// TIA Portal project "MoreLanguages" (V21)

(* hardware
DEVICE "PLC_Classic"  S7-300 station
   slot 0: "Rail_0"  Rail  6ES7 390-1***0-0AA0
   slot 2: "PLC_Classic"  CPU 315-2 PN/DP  6ES7 315-2EH14-0AB0  V3.2.18
      slot 2: "PROFINET interface_1"  PN-IO
         slot 1: "Port_1"  Port
         slot 2: "Port_2"  Port
DEVICE "PLC_More"  S7-1500 station
   slot 0: "Rail_0"  Rack  6ES7 590-1***0-0AA0
   slot 1: "PLC_More"  CPU 1516-3 PN/DP  6ES7 516-3AN02-0AB0  V2.9
      slot 3: "CPU display_1"  6ES7591-1BA00-0AA0
      slot 32768: "PROFINET interface_1"  X1
         slot 32769: "Port_1"  X1 P1
         slot 32770: "Port_2"  X1 P2
      slot 33024: "PROFINET interface_2"  X2
         slot 33025: "Port_1"  X2 P1
      slot 33280: "DP interface_1"  X3
      slot 34817: "Virtual CP interface port_1"  Virtual CP interface port  Virtual CP interface port
*)

// ===== PLC "PLC_Classic"  CPU 315-2 PN/DP =====

VAR_GLOBAL   // PLC tag table "Default tag table"
   "Tag__639308646888752274" AT %T1 : Timer;
   "Tag__639308646889222918" AT %I0.2 : Bool;
   "Tag__639308646889222919" AT %C1 : Counter;
   "Tag__639308646889222920" AT %I0.3 : Bool;
   "Tag__639308646889546626" AT %MW10 : Word;
   "Tag__639308646889705153" AT %QW0 : Word;
END_VAR

VAR_GLOBAL   // PLC tag table "IO"
   "Start" AT %I0.0 : Bool;   // Start button
   "Stop" AT %I0.1 : Bool;   // Stop button
   "Motor" AT %Q0.0 : Bool;   // Motor contactor
   "Raw" AT %IW2 : Int;   // Raw level
END_VAR

TYPE "Recipe"
   STRUCT
      amount : Int := 10;   // Units per batch
      heat : Bool;   // Whether the batch is heated
      dwell : Time := T#5S;   // Time in the heater
   END_STRUCT;
END_TYPE

DATA_BLOCK "Store"   // DB1
TITLE = Shared data
{ S7_Optimized_Access := 'FALSE' }
VERSION : 0.1
// A shared data block of a classic CPU, which has standard access only.
   VAR
      count : Int := 3;   // Batches made
      level : Word;
      current : "Recipe";
      flags : Array[0..7] of Bool;
   END_VAR
BEGIN
   current.amount := 12;
END_DATA_BLOCK

DATA_BLOCK "ScaleDb"   // DB2
{ S7_Optimized_Access := 'FALSE' }
VERSION : 0.1
// stored: InstanceOfName Scale
"Scale"
BEGIN
END_DATA_BLOCK

FUNCTION_BLOCK "Scale"   // FB1, SCL
TITLE = Scale a raw value
{ S7_Optimized_Access := 'FALSE' }
VERSION : 0.1
// SCL on a classic CPU.
   VAR_INPUT
      raw : Int;
      low : Real;
      high : Real;
   END_VAR
   VAR_OUTPUT
      value : Real;
   END_VAR
   VAR
      last : Real;
   END_VAR
BEGIN

    #value := #low + (#high - #low) * INT_TO_REAL(#raw) / 27648.0;
    #last := #value;
END_FUNCTION_BLOCK

FUNCTION_BLOCK "ClassicLad"   // FB10, LAD
TITLE = ClassicLad
{ S7_Optimized_Access := 'FALSE' }
// Ladder on a classic CPU, with global tags.
   VAR_INPUT
      enable : Bool;
   END_VAR
   VAR_OUTPUT
      running : Bool;
   END_VAR
   VAR
      latched : Bool;
   END_VAR
BEGIN

REGION Network 1: Run the motor
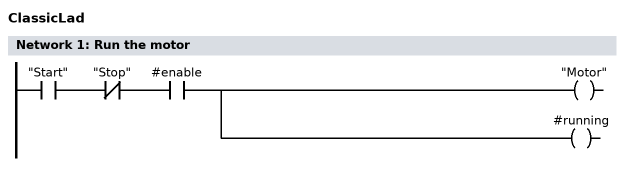
   RUNG wire#powerrail
      Contact( "Start" )
      I_Contact( "Stop" )
      Contact( #enable )
      wire#w1
      Coil( "Motor" )
   END_RUNG
   RUNG wire#w1
      Coil( #running )
   END_RUNG
   // the same network as SCL:
   "Motor" := "Start" AND NOT "Stop" AND #enable;
   #running := "Motor";
END_REGION
END_FUNCTION_BLOCK

FUNCTION_BLOCK "ClassicFbd"   // FB11, FBD
TITLE = ClassicFbd
{ S7_Optimized_Access := 'FALSE' }
// Function block diagram on a classic CPU.
   VAR_INPUT
      enable : Bool;
   END_VAR
   VAR_OUTPUT
      running : Bool;
   END_VAR
   VAR
      latched : Bool;
   END_VAR
BEGIN

REGION Network 1: Latch
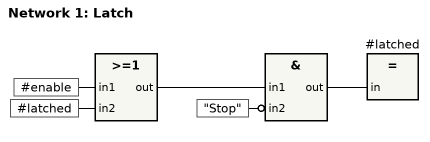
   #latched := (#enable OR #latched) AND NOT "Stop";
END_REGION
END_FUNCTION_BLOCK

FUNCTION "Classic" : Void   // FC1, STL
TITLE = Classic statement list
{ S7_Optimized_Access := 'FALSE' }
VERSION : 0.1
// An S5 timer, a counter, absolute addresses and a data block opened by number.
   VAR_INPUT
      start : Bool;
   END_VAR
   VAR_OUTPUT
      elapsed : Bool;
      parts : Word;
   END_VAR
BEGIN

REGION Network 1: An on-delay timer
         A     #start;
         L     S5T#2S;
         SD    "Tag__639308646888752274";
         A     "Tag__639308646888752274";
         =     #elapsed;
END_REGION

REGION Network 2: A counter
         A     "Tag__639308646889222918";
         CU    "Tag__639308646889222919";
         A     "Tag__639308646889222920";
         R     "Tag__639308646889222919";
         L     "Tag__639308646889222919";
         T     #parts;
END_REGION

REGION Network 3: A data block by number
         OPN   "Store";
         L     %DataW2;
         T     "Tag__639308646889546626";
         L     "Store".count;
         T     "Tag__639308646889705153";
END_REGION
END_FUNCTION

// ===== PLC "PLC_More"  CPU 1516-3 PN/DP =====

VAR_GLOBAL   // PLC tag table "Default tag table"
   "Tag__639308646937849854" AT %MD24 : DWord;
END_VAR

VAR_GLOBAL   // PLC tag table "IO"
   "Go" AT %I0.0 : Bool;   // Carriage start
   "Jammed" AT %I0.1 : Bool;   // Carriage jammed
   "Brake" AT %Q0.0 : Bool;   // Carriage brake
   "Pointer" AT %MD20 : DWord;   // Pointer for indirect access
END_VAR

// folder: Diagnosis

TYPE "Motor"
// A motor, assigned to a ProDiag function block where it is used.
   STRUCT
      running : Bool;
      tripped : Bool;
      ready : Bool;
      speed : Int;
   END_STRUCT;
END_TYPE

// folder: Common

DATA_BLOCK "BlinkDb"   // DB1
{ S7_Optimized_Access := 'TRUE' }
VERSION : 0.1
// stored: InstanceOfName Blink
"Blink"
BEGIN
END_DATA_BLOCK

// folder: Diagnosis

DATA_BLOCK "Plant"   // DB41
{ S7_Optimized_Access := 'TRUE' }
// Motors supervised by PlantDiag.
   VAR
      pump : "Motor";
      fans : Array[0..1] of "Motor";
      count : Int;
   END_VAR
BEGIN
END_DATA_BLOCK

DATA_BLOCK "LineDb"   // DB43
{ S7_Optimized_Access := 'TRUE' }
VERSION : 0.1
// stored: InstanceOfName Line
"Line"
BEGIN
END_DATA_BLOCK

DATA_BLOCK "PlantDiagDb"   // DB44
{ S7_Optimized_Access := 'TRUE' }
VERSION : 0.1
// stored: InstanceOfName PlantDiag
"PlantDiag"
BEGIN
END_DATA_BLOCK

// folder: (top level)

ORGANIZATION_BLOCK "ProDiagOB"   // OB250, ProDiag_OB, ProgramCycle
TITLE = "Main Program Sweep (Cycle)"
{ S7_Optimized_Access := 'TRUE' }
VERSION : 0.1
   VAR_INPUT
      Initial_Call : Bool;   // Initial call of this OB
      Remanence : Bool;   // =True, if remanent data are available
   END_VAR
BEGIN

REGION Network 1
   CALL "PlantDiag", "PlantDiagDb";
END_REGION
END_ORGANIZATION_BLOCK

// folder: Common

FUNCTION_BLOCK "Blink"   // FB1, SCL
TITLE = Blinker
{ S7_Optimized_Access := 'TRUE' }
VERSION : 0.1
// Toggles its output on every call while enabled.
   VAR_INPUT
      enable : Bool;
   END_VAR
   VAR_OUTPUT
      q : Bool;
   END_VAR
BEGIN

    IF #enable THEN
        #q := NOT #q;
    ELSE
        #q := FALSE;
    END_IF;
END_FUNCTION_BLOCK

// folder: Diagnosis

FUNCTION_BLOCK "Line"   // FB3, SCL
TITLE = Line with a motor
{ S7_Optimized_Access := 'TRUE' }
VERSION : 0.1
// A motor of a PLC data type in its static data; its instance data block is assigned to a ProDiag function block.
   VAR_INPUT
      command : Bool;
   END_VAR
   VAR_OUTPUT
      running : Bool;
   END_VAR
   VAR
      drive : "Motor";
   END_VAR
BEGIN

    #drive.running := #command AND #drive.ready AND NOT #drive.tripped;
    #running := #drive.running;
END_FUNCTION_BLOCK

FUNCTION_BLOCK "PlantDiag"   // FB42, ProDiag
{ S7_Optimized_Access := 'TRUE' }
   VAR
      PC_Flags : PC_Flags_V2;
      State : SV_FB_State_V2;
   END_VAR
   VAR_TEMP
      t_TempSvStateUDT : SV_State_V2;
      t_TempAlarmInstance : <type 200004f>;
      t_TempAsocValue1 : Variant;
      t_TempAsocValue2 : Variant;
      t_TempAsocValue3 : Variant;
   END_VAR
BEGIN
END_FUNCTION_BLOCK

// folder: Sequence

FUNCTION_BLOCK "Timed"   // FB30, GRAPH_PLUS
TITLE = Timed carriage
{ S7_Optimized_Access := 'TRUE' }
// A carriage that runs and brakes, with step times: the defaults, both set, and only the maximum set.
   VAR_INPUT
      ACK_EF : Bool := false;   // Acknowledge all errors and faults
      go : Bool;
      arrived : Bool;
      stopped : Bool;
      jammed : Bool;
   END_VAR
   VAR_OUTPUT
      motor : Bool;
      brake : Bool;
   END_VAR
   VAR
      HMI_INFO : Array[0..8] of UInt;
      IF_PAR : G7_IfParPlus_V6;
      RT_DATA : G7_RTDataPlus_V6;   // Internal data area
      Departs : G7_TransitionPlus_V6;   // Transition structure
      Reaches : G7_TransitionPlus_V6;   // Transition structure
      Rests : G7_TransitionPlus_V6;   // Transition structure
      Waiting : G7_StepPlus_V6;   // Step structure
      Running : G7_StepPlus_V6;   // Step structure
      Braking : G7_StepPlus_V6;   // Step structure
      SINI : Array[0..1] of USInt;
      LSTT : Array[0..2] of USInt;
      ATAJ : Array[0..2] of USInt;
      ATAB : Array[0..2] of USInt;
      PSTT : Array[0..2] of USInt;
      NSTT : Array[0..2] of USInt;
      ASSJ : Array[0..2] of USInt;
      ASSB : Array[0..2] of USInt;
      PTTS : Array[0..2] of USInt;
      NTTS : Array[0..2] of USInt;
      SW_SQTS : Array[0..2] of USInt;
      SWITCH : Array[0..0] of USInt;
      TVX : Array[0..1] of USInt;
      TTX : Array[0..1] of USInt;
      TSX : Array[0..1] of USInt;
      S00X : Array[0..1] of USInt;
      SOFFX : Array[0..1] of USInt;
      SONX : Array[0..1] of USInt;
      SAX : Array[0..1] of USInt;
      SERRX : Array[0..3] of USInt;
      SMX : Array[0..3] of USInt;
      S0X : Array[0..3] of USInt;
      S1X : Array[0..3] of USInt;
      IL_ALARM_INST : Diag_Alarm;
      SUP_ALARM_INST : Diag_Alarm;
      STEP_TIME_ALARM_INST : Diag_Alarm;
      IEC_TIMER_INST : IEC_TIMER;
      TRANSACTION_FLAG : Bool := false;
   END_VAR
   // SINI[0] := 2;
   // LSTT[0] := 255;
   // LSTT[1] := 255;
   // ATAJ[1] := 1;
   // ATAJ[2] := 2;
   // ATAB[1] := 1;
   // ATAB[2] := 2;
   // PSTT[1] := 1;
   // PSTT[2] := 2;
   // NSTT[0] := 1;
   // NSTT[1] := 2;
   // ASSJ[1] := 1;
   // ASSJ[2] := 2;
   // ASSB[1] := 1;
   // ASSB[2] := 2;
   // PTTS[0] := 255;
   // PTTS[2] := 1;
   // NTTS[1] := 1;
   // NTTS[2] := 2;
   // TVX[0] := 16#1;
   // TTX[0] := 16#1;
   // TSX[0] := 16#1;
   // S00X[0] := 16#1;
   // SOFFX[0] := 16#1;
   // SONX[0] := 16#1;
   // SAX[0] := 16#1;
   // SERRX[0] := 16#1;
   // SMX[0] := 16#1;
   // S0X[0] := 16#1;
   // S1X[0] := 16#1;
BEGIN
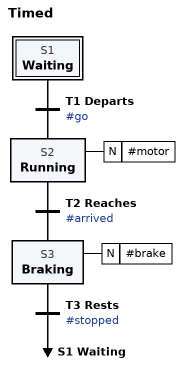
   // sequencer 1
   INITIAL_STEP Waiting:   // S1, max time T#10S, warning time T#7S
   END_STEP
   TRANSITION Departs FROM Waiting TO Running   // T1
      := #go;
   END_TRANSITION
   STEP Running:   // S2, max time T#30S, warning time T#20S
      supervision V := #jammed;
              N    #motor
   END_STEP
   TRANSITION Reaches FROM Running TO Braking   // T2
      := #arrived;
   END_TRANSITION
   STEP Braking:   // S3, max time T#1M30S, warning time T#7S
              N    #brake
   END_STEP
   TRANSITION Rests FROM Braking TO Waiting   // T3, jump
      := #stopped;
   END_TRANSITION
END_FUNCTION_BLOCK

// folder: Statement

FUNCTION_BLOCK "StlForms"   // FB2, STL
TITLE = More statement list
{ S7_Optimized_Access := 'TRUE' }
VERSION : 0.1
// Word logic, shifts, conversions, a jump list, a loop, status bits, edges, constants and calls of function blocks.
   VAR_INPUT
      mode : Int;
      raw : Word;
      count : Int;
      start : Bool;
   END_VAR
   VAR_OUTPUT
      result : DInt;
      ratio : Real;
      done : Bool;
      blinking : Bool;
   END_VAR
   VAR
      rising : Bool;
      falling : Bool;
      blinker : "Blink";
   END_VAR
   VAR_TEMP
      w : Word;
      d : DWord;
      i : Int;
      loops : Int;
      duration : Time;
      s5 : S5Time;
      "b" : Byte;
      ch : Char;
   END_VAR
BEGIN

REGION Network 1: Word logic
         L     #raw;
         AW    W#16#FF00;
         OW    W#16#000F;
         XOW   W#16#0101;
         INVI;
         T     #w;
END_REGION

REGION Network 2: Shifts and rotates
         L     #raw;
         SLW   2;
         SRW   1;
         T     #w;
         L     #count;
         SSI   3;
         T     #i;
         L     DW#16#8000_0001;
         RLD   1;
         RRD   2;
         T     #d;
END_REGION

REGION Network 3: Conversions
         L     #count;
         ITD;
         DTR;
         T     #ratio;
         RND;
         T     #result;
         L     #ratio;
         TRUNC;
         T     #result;
         L     #count;
         ITB;
         T     #w;
         BTI;
         T     #i;
END_REGION

REGION Network 4: A jump list
         L     #mode;
         JL    over;
         JU    zero;
         JU    one;
   over: JU    fin;
   zero: L     0;
         JU    keep;
   one:  L     1;
   keep: T     #i;
   fin:  NOP   0;
END_REGION

REGION Network 5: A loop
         L     0;
         T     #i;
         L     5;
   next: T     #loops;
         L     #i;
         +     1;
         T     #i;
         L     #loops;
         LOOP  next;
END_REGION

REGION Network 6: Status bits
         L     #count;
         L     1000;
         *I;
         T     #i;
         A     OV;
         =     #done;
         SET;
         SAVE;
         CLR;
         A     BR;
         NOT;
         =     #done;
END_REGION

REGION Network 7: Edges, set and reset
         A     #start;
         FP    #rising;
         S     #done;
         A     #start;
         FN    #falling;
         R     #done;
END_REGION

REGION Network 8: Constants
         L     2#1010_1010;
         T     #"b";
         L     B#16#1F;
         T     #"b";
         L     W#16#1F2E;
         T     #w;
         L     1500.0;
         T     #ratio;
         L     T#1S500MS;
         T     #duration;
         L     S5T#2S;
         T     #s5;
         L     'AB';
         T     #w;
         L     'A';
         T     #ch;
         L     DINT#100000;
         T     #result;
         L     C#100;
         T     #w;
END_REGION

REGION Network 9: Calls of function blocks
         CALL  "Blink", "BlinkDb"
         ( enable := #start,
           q      :=
         );
         CALL  #blinker
         ( enable := #done,
           q      := #blinking
         );
END_REGION

REGION Network 10: A conditional end
         A     #done;
         BEC;
         L     0;
         T     #i;
END_REGION
END_FUNCTION_BLOCK

FUNCTION "StlIndirect" : Void   // FC1, STL
TITLE = Indirect addressing
{ S7_Optimized_Access := 'FALSE' }
VERSION : 0.1
// Pointers in a variable and in the address registers, which need a block with standard access.
   VAR_INPUT
      index : Int;
      dbNo : Int;
   END_VAR
   VAR_OUTPUT
      value : Int;
      flag : Bool;
      address : DWord;
   END_VAR
   VAR_TEMP
      place : DWord;
      dbNumber : Word;
      local : Array[0..3] of Int;
   END_VAR
BEGIN

REGION Network 1: Memory-indirect, through a pointer in a variable
   // The index counts bytes; shifting it by three makes it a bit address.
         L     #index;
         SLD   3;
         T     #place;
         L     MW[#place];
         T     #value;
         A     I[#place];
         =     #flag;
END_REGION

REGION Network 2: Register-indirect within an area
         L     P#10.0;
         LAR1;
         L     MW[AR1,P#2.0];
         T     #value;
         +AR1  P#4.0;
         A     M[AR1,P#0.1];
         =     #flag;
         TAR1  "Tag__639308646937849854";
END_REGION

REGION Network 3: Register-indirect across areas
         L;
         LAR1;
         L     W[AR1,P#2.0];  // the second element
         T     #value;
         LAR2  P#M20.0;
         A     [AR2,P#0.1];
         =     #flag;
         TAR2;
         T     #address;
END_REGION

REGION Network 4: A data block opened through a variable
         L     #dbNo;
         T     #dbNumber;
         OPN   DB[#dbNumber];
         L     DBW[AR1,P#0.0];
         T     #value;
         L     DBNO;
         L     DBLG;
         CAR;
END_REGION
END_FUNCTION